FUNCTION_BLOCK basicForcaDO (* Forcamento de saidas digitais pela IHM: saida = comando da logica ou valor forcado (LIGADO/DESLIGADO) *)
  (* Standard: 61499-2 *)
  (* Version 1.0, 20/10/2026, Hidryco, Hidryco, 1.0: criado para o IO_DQ32 (forcamento por bit no simbolo) *)
  PACKAGE Hidryco.HidrycoLib;
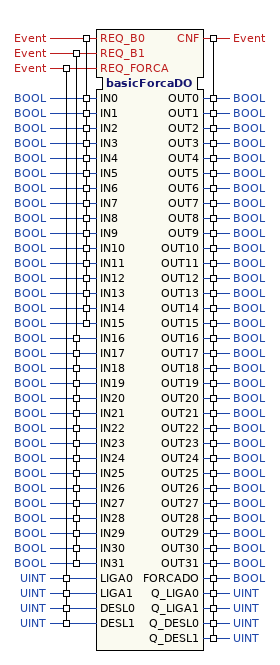
  EVENT_INPUT
    REQ_B0 WITH IN0, IN1, IN2, IN3, IN4, IN5, IN6, IN7, IN8, IN9, IN10, IN11, IN12, IN13, IN14, IN15; (* Novos comandos dos bits 0-15 *)
    REQ_B1 WITH IN16, IN17, IN18, IN19, IN20, IN21, IN22, IN23, IN24, IN25, IN26, IN27, IN28, IN29, IN30, IN31; (* Novos comandos dos bits 16-31 *)
    REQ_FORCA WITH LIGA0, LIGA1, DESL0, DESL1; (* Novas mascaras de forcamento (IHM) *)
  END_EVENT
  EVENT_OUTPUT
    CNF WITH OUT0, OUT1, OUT2, OUT3, OUT4, OUT5, OUT6, OUT7, OUT8, OUT9, OUT10, OUT11, OUT12, OUT13, OUT14, OUT15, OUT16, OUT17, OUT18, OUT19, OUT20, OUT21, OUT22, OUT23, OUT24, OUT25, OUT26, OUT27, OUT28, OUT29, OUT30, OUT31, FORCADO, Q_LIGA0, Q_LIGA1, Q_DESL0, Q_DESL1; (* Saidas efetivas atualizadas *)
  END_EVENT
  VAR_INPUT
    IN0 : BOOL; (* Comando do bit 0 (logica) *)
    IN1 : BOOL; (* Comando do bit 1 (logica) *)
    IN2 : BOOL; (* Comando do bit 2 (logica) *)
    IN3 : BOOL; (* Comando do bit 3 (logica) *)
    IN4 : BOOL; (* Comando do bit 4 (logica) *)
    IN5 : BOOL; (* Comando do bit 5 (logica) *)
    IN6 : BOOL; (* Comando do bit 6 (logica) *)
    IN7 : BOOL; (* Comando do bit 7 (logica) *)
    IN8 : BOOL; (* Comando do bit 8 (logica) *)
    IN9 : BOOL; (* Comando do bit 9 (logica) *)
    IN10 : BOOL; (* Comando do bit 10 (logica) *)
    IN11 : BOOL; (* Comando do bit 11 (logica) *)
    IN12 : BOOL; (* Comando do bit 12 (logica) *)
    IN13 : BOOL; (* Comando do bit 13 (logica) *)
    IN14 : BOOL; (* Comando do bit 14 (logica) *)
    IN15 : BOOL; (* Comando do bit 15 (logica) *)
    IN16 : BOOL; (* Comando do bit 16 (logica) *)
    IN17 : BOOL; (* Comando do bit 17 (logica) *)
    IN18 : BOOL; (* Comando do bit 18 (logica) *)
    IN19 : BOOL; (* Comando do bit 19 (logica) *)
    IN20 : BOOL; (* Comando do bit 20 (logica) *)
    IN21 : BOOL; (* Comando do bit 21 (logica) *)
    IN22 : BOOL; (* Comando do bit 22 (logica) *)
    IN23 : BOOL; (* Comando do bit 23 (logica) *)
    IN24 : BOOL; (* Comando do bit 24 (logica) *)
    IN25 : BOOL; (* Comando do bit 25 (logica) *)
    IN26 : BOOL; (* Comando do bit 26 (logica) *)
    IN27 : BOOL; (* Comando do bit 27 (logica) *)
    IN28 : BOOL; (* Comando do bit 28 (logica) *)
    IN29 : BOOL; (* Comando do bit 29 (logica) *)
    IN30 : BOOL; (* Comando do bit 30 (logica) *)
    IN31 : BOOL; (* Comando do bit 31 (logica) *)
    LIGA0 : UINT; (* Forcar LIGADO: mascara dos bits 0-15 (bit k = saida k) *)
    LIGA1 : UINT; (* Forcar LIGADO: mascara dos bits 16-31 (bit k = saida 16+k) *)
    DESL0 : UINT; (* Forcar DESLIGADO: mascara dos bits 0-15 *)
    DESL1 : UINT; (* Forcar DESLIGADO: mascara dos bits 16-31 *)
  END_VAR
  VAR_OUTPUT
    OUT0 : BOOL; (* Saida efetiva do bit 0 (comando ou forcamento) *)
    OUT1 : BOOL; (* Saida efetiva do bit 1 (comando ou forcamento) *)
    OUT2 : BOOL; (* Saida efetiva do bit 2 (comando ou forcamento) *)
    OUT3 : BOOL; (* Saida efetiva do bit 3 (comando ou forcamento) *)
    OUT4 : BOOL; (* Saida efetiva do bit 4 (comando ou forcamento) *)
    OUT5 : BOOL; (* Saida efetiva do bit 5 (comando ou forcamento) *)
    OUT6 : BOOL; (* Saida efetiva do bit 6 (comando ou forcamento) *)
    OUT7 : BOOL; (* Saida efetiva do bit 7 (comando ou forcamento) *)
    OUT8 : BOOL; (* Saida efetiva do bit 8 (comando ou forcamento) *)
    OUT9 : BOOL; (* Saida efetiva do bit 9 (comando ou forcamento) *)
    OUT10 : BOOL; (* Saida efetiva do bit 10 (comando ou forcamento) *)
    OUT11 : BOOL; (* Saida efetiva do bit 11 (comando ou forcamento) *)
    OUT12 : BOOL; (* Saida efetiva do bit 12 (comando ou forcamento) *)
    OUT13 : BOOL; (* Saida efetiva do bit 13 (comando ou forcamento) *)
    OUT14 : BOOL; (* Saida efetiva do bit 14 (comando ou forcamento) *)
    OUT15 : BOOL; (* Saida efetiva do bit 15 (comando ou forcamento) *)
    OUT16 : BOOL; (* Saida efetiva do bit 16 (comando ou forcamento) *)
    OUT17 : BOOL; (* Saida efetiva do bit 17 (comando ou forcamento) *)
    OUT18 : BOOL; (* Saida efetiva do bit 18 (comando ou forcamento) *)
    OUT19 : BOOL; (* Saida efetiva do bit 19 (comando ou forcamento) *)
    OUT20 : BOOL; (* Saida efetiva do bit 20 (comando ou forcamento) *)
    OUT21 : BOOL; (* Saida efetiva do bit 21 (comando ou forcamento) *)
    OUT22 : BOOL; (* Saida efetiva do bit 22 (comando ou forcamento) *)
    OUT23 : BOOL; (* Saida efetiva do bit 23 (comando ou forcamento) *)
    OUT24 : BOOL; (* Saida efetiva do bit 24 (comando ou forcamento) *)
    OUT25 : BOOL; (* Saida efetiva do bit 25 (comando ou forcamento) *)
    OUT26 : BOOL; (* Saida efetiva do bit 26 (comando ou forcamento) *)
    OUT27 : BOOL; (* Saida efetiva do bit 27 (comando ou forcamento) *)
    OUT28 : BOOL; (* Saida efetiva do bit 28 (comando ou forcamento) *)
    OUT29 : BOOL; (* Saida efetiva do bit 29 (comando ou forcamento) *)
    OUT30 : BOOL; (* Saida efetiva do bit 30 (comando ou forcamento) *)
    OUT31 : BOOL; (* Saida efetiva do bit 31 (comando ou forcamento) *)
    FORCADO : BOOL; (* Alguma saida do cartao forcada *)
    Q_LIGA0 : UINT; (* Mascara LIGA0 em uso (para a IHM) *)
    Q_LIGA1 : UINT; (* Mascara LIGA1 em uso (para a IHM) *)
    Q_DESL0 : UINT; (* Mascara DESL0 em uso (para a IHM) *)
    Q_DESL1 : UINT; (* Mascara DESL1 em uso (para a IHM) *)
  END_VAR
  VAR
    wL0 : WORD;
    wL1 : WORD;
    wD0 : WORD;
    wD1 : WORD;
  END_VAR
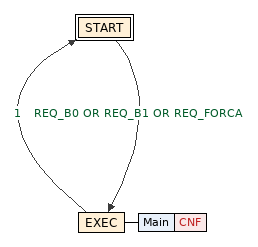
  EC_STATES
    START; (* Initial State *)
    EXEC : Main -> CNF;
  END_STATES
  EC_TRANSITIONS
    START TO EXEC := REQ_B0 OR REQ_B1 OR REQ_FORCA;
    EXEC TO START := 1;
  END_TRANSITIONS
  ALGORITHM Main IN ST: (* Aplica o forcamento *)
(* Saida efetiva = comando da logica, a nao ser que o bit esteja forcado pela IHM.
   LIGAx: bit em 1 = saida forcada LIGADA; DESLx: bit em 1 = saida forcada DESLIGADA (DESL prevalece).
   Mascaras nao sao persistentes: depois de reiniciar o CLP nenhuma saida fica forcada. *)
wL0 := UINT_TO_WORD(LIGA0); wL1 := UINT_TO_WORD(LIGA1);
wD0 := UINT_TO_WORD(DESL0); wD1 := UINT_TO_WORD(DESL1);
OUT0 := (IN0 OR ((wL0 AND 16#0001) <> 0)) AND ((wD0 AND 16#0001) = 0);
OUT1 := (IN1 OR ((wL0 AND 16#0002) <> 0)) AND ((wD0 AND 16#0002) = 0);
OUT2 := (IN2 OR ((wL0 AND 16#0004) <> 0)) AND ((wD0 AND 16#0004) = 0);
OUT3 := (IN3 OR ((wL0 AND 16#0008) <> 0)) AND ((wD0 AND 16#0008) = 0);
OUT4 := (IN4 OR ((wL0 AND 16#0010) <> 0)) AND ((wD0 AND 16#0010) = 0);
OUT5 := (IN5 OR ((wL0 AND 16#0020) <> 0)) AND ((wD0 AND 16#0020) = 0);
OUT6 := (IN6 OR ((wL0 AND 16#0040) <> 0)) AND ((wD0 AND 16#0040) = 0);
OUT7 := (IN7 OR ((wL0 AND 16#0080) <> 0)) AND ((wD0 AND 16#0080) = 0);
OUT8 := (IN8 OR ((wL0 AND 16#0100) <> 0)) AND ((wD0 AND 16#0100) = 0);
OUT9 := (IN9 OR ((wL0 AND 16#0200) <> 0)) AND ((wD0 AND 16#0200) = 0);
OUT10 := (IN10 OR ((wL0 AND 16#0400) <> 0)) AND ((wD0 AND 16#0400) = 0);
OUT11 := (IN11 OR ((wL0 AND 16#0800) <> 0)) AND ((wD0 AND 16#0800) = 0);
OUT12 := (IN12 OR ((wL0 AND 16#1000) <> 0)) AND ((wD0 AND 16#1000) = 0);
OUT13 := (IN13 OR ((wL0 AND 16#2000) <> 0)) AND ((wD0 AND 16#2000) = 0);
OUT14 := (IN14 OR ((wL0 AND 16#4000) <> 0)) AND ((wD0 AND 16#4000) = 0);
OUT15 := (IN15 OR ((wL0 AND 16#8000) <> 0)) AND ((wD0 AND 16#8000) = 0);
OUT16 := (IN16 OR ((wL1 AND 16#0001) <> 0)) AND ((wD1 AND 16#0001) = 0);
OUT17 := (IN17 OR ((wL1 AND 16#0002) <> 0)) AND ((wD1 AND 16#0002) = 0);
OUT18 := (IN18 OR ((wL1 AND 16#0004) <> 0)) AND ((wD1 AND 16#0004) = 0);
OUT19 := (IN19 OR ((wL1 AND 16#0008) <> 0)) AND ((wD1 AND 16#0008) = 0);
OUT20 := (IN20 OR ((wL1 AND 16#0010) <> 0)) AND ((wD1 AND 16#0010) = 0);
OUT21 := (IN21 OR ((wL1 AND 16#0020) <> 0)) AND ((wD1 AND 16#0020) = 0);
OUT22 := (IN22 OR ((wL1 AND 16#0040) <> 0)) AND ((wD1 AND 16#0040) = 0);
OUT23 := (IN23 OR ((wL1 AND 16#0080) <> 0)) AND ((wD1 AND 16#0080) = 0);
OUT24 := (IN24 OR ((wL1 AND 16#0100) <> 0)) AND ((wD1 AND 16#0100) = 0);
OUT25 := (IN25 OR ((wL1 AND 16#0200) <> 0)) AND ((wD1 AND 16#0200) = 0);
OUT26 := (IN26 OR ((wL1 AND 16#0400) <> 0)) AND ((wD1 AND 16#0400) = 0);
OUT27 := (IN27 OR ((wL1 AND 16#0800) <> 0)) AND ((wD1 AND 16#0800) = 0);
OUT28 := (IN28 OR ((wL1 AND 16#1000) <> 0)) AND ((wD1 AND 16#1000) = 0);
OUT29 := (IN29 OR ((wL1 AND 16#2000) <> 0)) AND ((wD1 AND 16#2000) = 0);
OUT30 := (IN30 OR ((wL1 AND 16#4000) <> 0)) AND ((wD1 AND 16#4000) = 0);
OUT31 := (IN31 OR ((wL1 AND 16#8000) <> 0)) AND ((wD1 AND 16#8000) = 0);
FORCADO := (LIGA0 <> 0) OR (LIGA1 <> 0) OR (DESL0 <> 0) OR (DESL1 <> 0);
Q_LIGA0 := LIGA0; Q_LIGA1 := LIGA1; Q_DESL0 := DESL0; Q_DESL1 := DESL1;
  END_ALGORITHM
END_FUNCTION_BLOCK
